(* IEC 61131-3 sources: Lasal-MCP/examples/SampleSource/LASALScreenAdvancedSolution/LASALScreenAdvancedSolution/LASALScreenAdvacnedSolution/Stations/Terminal/HMI/Network/GlobalNet, 1 file *)

(* ---- ONE_GlobalNet_Table.st ---- *)
#define OBJECTS_CONFIG

FUNCTION GLOBAL TAB ONE_GlobalNet
-1$UINT, 0$UINT,
0$UINT, 0$UINT,

4$UDINT,
TO_UDINT(3788417926), "_Global", 0$UINT, 15$UINT, 0$UINT,
TO_UDINT(1683757165), "MyKeyboardCode", 0$UINT, 0$UINT, 1$UINT,
TO_UDINT(2348910643), "MyRecalculate", 0$UINT, 0$UINT, 1$UINT,
TO_UDINT(2682062625), "MyUserCall", 0$UINT, 0$UINT, 1$UINT,

_NO_ATTR, TO_UDINT(2965089866), "MYKEYBOARDCODE1",

_NO_ATTR, TO_UDINT(1015058217), "MYRECALCULATE1",

_NO_ATTR, TO_UDINT(3475645166), "MYUSERCALL1",

//Internal connections
0$UDINT,
0$UDINT,
0$UDINT,
0$UDINT,

//Initialization values
0$UDINT,
0$UDINT,

//Symbolic initialization values
0$UDINT,
0$UDINT,

//Initialization of string values
0$UDINT,
0$UDINT,

//Configuration of tasks (RealTime, Cyclic, Background)
0$UDINT,
0$UDINT,

0$UDINT,
0$UDINT,

0$UDINT,
0$UDINT,

//External connections
0$UDINT,
3$UDINT,
TO_UDINT(0), "Lse", C_DIR, TO_UDINT(299963966), "Lse","Lse",
TO_UDINT(1), "Lse", C_DIR, TO_UDINT(299963966), "Lse","Lse",
TO_UDINT(2), "Lse", C_DIR, TO_UDINT(299963966), "Lse","Lse",

//Magic internal connections
0$UDINT,
0$UDINT,

//Configuration of timeslots of tasks (RealTime, Cyclic)
#ifdef __LSLLDR_TIMESLOTS__
0$UDINT,
0$UDINT,

0$UDINT,
0$UDINT,

#endif //__LSLLDR_TIMESLOTS__

//MultiMaster connections
#ifdef __LSLLDR_MULTIMASTER__
0$UDINT,
0$UDINT,
#endif //__LSLLDR_MULTIMASTER__

//Configuration for task ID (RealTime, CyclicTime)
#ifdef __LSLLDR_TASKID__
"\\\\TASKS2  "
0$UDINT,
0$UDINT,

0$UDINT,
0$UDINT,

0$UDINT,
0$UDINT,

#endif //__LSLLDR_TASKID__

END_FUNCTION
